// TIA Portal V20 export
// export: Created 2026-10-22T17:35:50.4361467Z, ExportSetting WithDefaults
ORGANIZATION_BLOCK "Main"   // OB1, LAD, ProgramCycle
TITLE = Main program sweep (cycle)
{ S7_Optimized_Access := 'TRUE' }
VERSION : 0.1
// stored: AutoNumber true, IsIECCheckEnabled true, SetENOAutomatically false
   VAR_INPUT
      Initial_Call : Bool;   // Initial call of this OB
   END_VAR
   VAR_TEMP
      start : Bool;
      stop : Bool;
      latch : Bool;   // Motor latched on
      count : Int;
      big : Bool;
      delayed : Bool;
      "a" : Bool;
      "b" : Bool;
      text : String;
   END_VAR
   VAR_TEMP   // added for the SCL form of the ladder/FBD networks
      _w1 : Bool;
   END_VAR
BEGIN

REGION Network 1: Seal-in
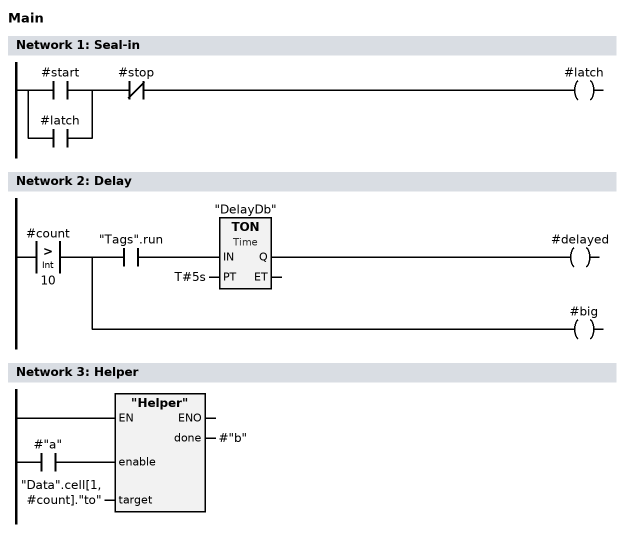
   RUNG wire#powerrail
      Contact( #start )
      wire#w1
      I_Contact( #stop )
      Coil( #latch )
   END_RUNG
   RUNG wire#powerrail
      Contact( #latch )
   END_RUNG wire#w1
   // the same network as SCL:
   #latch := (#start OR #latch) AND NOT #stop;
END_REGION

REGION Network 2: Delay
   RUNG wire#powerrail
      { S7_Templates := "SrcType := Int" } GT_Contact(in1 := #count, in2 := 10)
      wire#w1
      Contact( "Tags".run )
      { S7_Templates := "time_type := Time" } "DelayDb".TON(pt := T#5s, et =>)
      Coil( #delayed )
   END_RUNG
   RUNG wire#w1
      Coil( #big )
   END_RUNG
   // the same network as SCL:
   #_w1 := #count > 10;
   "DelayDb".TON(IN := #_w1 AND "Tags".run, PT := T#5s);
   #delayed := "DelayDb".Q;
   #big := #_w1;
END_REGION

REGION Network 3: Helper
   RUNG wire#powerrail
      "Helper"(enable := wire#w1, done => #"b", target := "Data".cell[1, #count]."to")
   END_RUNG
   RUNG wire#powerrail
      Contact( #"a" )
   END_RUNG wire#w1
   // the same network as SCL:
   "Helper"(enable := #"a", target := "Data".cell[1, #count]."to", done => #"b");
END_REGION

REGION Network 4 (SCL): Cell text
   // Text of the cell
   #text := CONCAT_STRING(IN1 := 'cell ', IN2 := "Data".to.name);
   #count := "Count"(#text);
END_REGION
END_ORGANIZATION_BLOCK
